// TIA Portal V21 export
// export: Created 2000-01-01T00:00:00.0000000Z, ExportSetting None
TYPE "UDT_HMI_FIO_Assembler"
   STRUCT
      bManualMode { ExternalWritable := 'False'} : Bool;   // TRUE手动, FALSE自动
      bStartCmd { ExternalWritable := 'False'} : Bool;   // HMI启动命令
      bStopCmd { ExternalWritable := 'False'} : Bool;   // HMI停止命令
      bResetCmd { ExternalWritable := 'False'} : Bool;   // HMI故障复位命令
      tActionDelay { ExternalWritable := 'False'} : Time;   // 气缸定位/夹紧保持延时（默认 T#500ms）
      tStepTimeout { ExternalWritable := 'False'} : Time;   // 单步动作超时时间（默认 T#6s）
      iCurrentStep { ExternalWritable := 'False'} : Int;   // 状态反馈：当前装配顺控步号
      diAssembledCount { ExternalWritable := 'False'} : DInt;   // 状态反馈：累计完成装配成品数
      bRunning { ExternalWritable := 'False'} : Bool;   // 状态反馈：运行中
      bFault { ExternalWritable := 'False'} : Bool;   // 状态反馈：超时或急停故障
      wStatus { ExternalWritable := 'False'} : Word;   // 状态码：16#0000正常, 16#7000待机, 16#8401工位超时, 16#8402急停触发
   END_STRUCT;
END_TYPE
